(* IEC 61131-3 sources: s7-to-codesys/tests/POUs/S7Compat/FB_F_ScaleX_Test, 9 files *)

(* ---- FB_F_ScaleX_Test.decl.st ---- *)
// Назначение: набор тестов CfUnit (coUnit 1.2.0.0) для F_ScaleX — аналога S7 SCALE_X:
//             середина и границы диапазона, VALUE ниже 0.0 и выше 1.0 (линейное
//             продолжение), диапазон с отрицательной границей, вырожденный и обратный
//             диапазон (та же формула). Ожидаемые значения — по формуле Siemens
//             OUT = VALUE * (MAX - MIN) + MIN, а не по результату реализации.
//             Экземпляр набора объявляется в PRG_Tests (объявление регистрирует набор).
// Автор:      kr0nsch
// Версия:     0.1.0
// Документ:   docs/MAPPING.md, раздел «NORM_X и SCALE_X»
FUNCTION_BLOCK FB_F_ScaleX_Test EXTENDS coUnit.FB_TestSuite
VAR CONSTANT
    // арифметика REAL: сравнение с допуском
    R_DELTA : REAL := 0.0001;
END_VAR

(* ---- AboveOneExtrapolates.method.decl.st ---- *)
// F_ScaleX(rMin := 0.0, rValue := 1.2, rMax := 100.0) = 120.0.
METHOD PRIVATE AboveOneExtrapolates
VAR
    rResult : REAL;     // результат F_ScaleX
END_VAR

(* ---- BelowZeroExtrapolates.method.decl.st ---- *)
// F_ScaleX(rMin := 0.0, rValue := -0.25, rMax := 100.0) = -25.0.
METHOD PRIVATE BelowZeroExtrapolates
VAR
    rResult : REAL;     // результат F_ScaleX
END_VAR

(* ---- EqualBoundsGivesMin.method.decl.st ---- *)
// F_ScaleX(rMin := 10.0, rValue := 0.5, rMax := 10.0) = 10.0.
METHOD PRIVATE EqualBoundsGivesMin
VAR
    rResult : REAL;     // результат F_ScaleX
END_VAR

(* ---- HalfGivesMidRange.method.decl.st ---- *)
// F_ScaleX(rMin := 0.0, rValue := 0.5, rMax := 100.0) = 50.0.
METHOD PRIVATE HalfGivesMidRange
VAR
    rResult : REAL;     // результат F_ScaleX
END_VAR

(* ---- NegativeLowBound.method.decl.st ---- *)
// F_ScaleX(rMin := -50.0, rValue := 0.75, rMax := 50.0) = 25.0.
METHOD PRIVATE NegativeLowBound
VAR
    rResult : REAL;     // результат F_ScaleX
END_VAR

(* ---- OneGivesMax.method.decl.st ---- *)
// F_ScaleX(rMin := 20.0, rValue := 1.0, rMax := 80.0) = 80.0.
METHOD PRIVATE OneGivesMax
VAR
    rResult : REAL;     // результат F_ScaleX
END_VAR

(* ---- ReversedBoundsKeepsFormula.method.decl.st ---- *)
// F_ScaleX(rMin := 100.0, rValue := 0.25, rMax := 0.0) = 75.0.
METHOD PRIVATE ReversedBoundsKeepsFormula
VAR
    rResult : REAL;     // результат F_ScaleX
END_VAR

(* ---- ZeroGivesMin.method.decl.st ---- *)
// F_ScaleX(rMin := 20.0, rValue := 0.0, rMax := 80.0) = 20.0.
METHOD PRIVATE ZeroGivesMin
VAR
    rResult : REAL;     // результат F_ScaleX
END_VAR
